Staubli VAL3: click_refreshRobotMsg.pgx

program click_refreshRobotMsg()
begin
  nMsgType=1
  call initMsg()
  call rs:getLog(sRobotMsg,nMsgType)
  userPageSet("message","btnAllMsg","style.backgroundColor","#FFFFFF")
  userPageSet("message","btnRobotMsg","style.backgroundColor","#33FF33")
  userPageSet("message","btnTrajMsg","style.backgroundColor","#FFFFFF")
  userPageSet("message","btnIOMsg","style.backgroundColor","#FFFFFF")
end
